(* IEC 61131-3 sources: nautilus/examples/lift-station/lib, 2 files *)

(* ---- physics.st ---- *)
(* Bench-only plant model: a wet-well level integrator and a submersible
   pump/VFD dynamic model. Two FUNCTION_BLOCKs, no PROGRAM — a project
   library (docs/functions.md "A .ld library", the same rule for .st).
   sim.st is the only caller; field.yaml has no sim task, so these two
   blocks sit compiled but unused in that manifest — harmless dead code,
   the same way a project's other library functions are. *)

FUNCTION_BLOCK WetWellModel
(* Integrates a level from an inflow/outflow balance. WW-101: a 13 ft
   level span over 1,320 gal of usable volume between the span's limits,
   so 13.2 gal per %: 100 gpm net moves the level 1 % in about 8 s. *)
VAR_INPUT
    InflowGpm  : REAL;
    OutflowGpm : REAL;
    Dt         : REAL; (* seconds *)
END_VAR
VAR_IN_OUT
    Level : REAL; (* %, 0..100 *)
END_VAR
VAR CONSTANT
    GalPerPercent : REAL := 13.2; (* 1,320 gal span / 100 % = 13.2 gal per % *)
END_VAR
(* gal/min * s / 60 = gal *)
Level := LIMIT(0.0, Level + (InflowGpm - OutflowGpm) * Dt / 60.0 / GalPerPercent, 100.0);
END_FUNCTION_BLOCK

FUNCTION_BLOCK VfdModel
(* A submersible pump + VFD, standing in for the field device on the
   bench: RunCmd/SpeedCmd in, Running/SpeedHz/Amps/Fault out. Running lags
   RunCmd by 0.5 s (starter contactor + soft-start), and drops the instant
   a fault is injected. SpeedHz ramps toward SpeedCmd at 10 Hz/s while
   commanded and running, and ramps back to 0 otherwise. Amps follows
   speed-squared, the affinity-law shape a centrifugal load actually
   draws. Fault is a plain pass-through of the bench inject tag — a real
   VFD's own fault relay, not the ladder's fail-to-run latch (that is a
   separate, higher-level condition computed in permissives.ld). *)
VAR_INPUT
    RunCmd      : BOOL;
    SpeedCmd    : REAL;
    Dt          : REAL;
    InjectFault : BOOL;
END_VAR
VAR_OUTPUT
    Running : BOOL;
    SpeedHz : REAL;
    Amps    : REAL;
    Fault   : BOOL;
END_VAR
VAR
    t1 : TON;
END_VAR
VAR CONSTANT
    RampHzPerS : REAL := 10.0; (* speed ramp rate *)
    FullLoadA  : REAL := 22.0; (* amps at MaxHz, full load *)
    MaxHz      : REAL := 60.0; (* VFD speed ceiling *)
END_VAR
Fault := InjectFault;
t1(IN := RunCmd AND NOT Fault, PT := T#500MS);
Running := t1.Q;
IF Running THEN
    SpeedHz := LIMIT(0.0, SpeedHz + LIMIT(-RampHzPerS * Dt, SpeedCmd - SpeedHz, RampHzPerS * Dt), MaxHz);
ELSE
    SpeedHz := MAX(0.0, SpeedHz - RampHzPerS * Dt);
END_IF;
Amps := (SpeedHz / MaxHz) * (SpeedHz / MaxHz) * FullLoadA;
END_FUNCTION_BLOCK

(* ---- pump.st ---- *)
(* Runtime accounting shared by both pumps: a retained UDT (PumpStats) and
   a FUNCTION_BLOCK that updates it by reference, so neither the sequence
   nor the permissives ever touch accumulation math themselves. A .st file
   with no PROGRAM is a project library — see docs/functions.md "A .ld
   library" (the same rule, one language over). *)

TYPE
  PumpStats : STRUCT
    Starts     : INT;   (* start count *)
    Hours      : REAL;  (* run hours *)
    LastRunSec : REAL;  (* length of the most recently completed run *)
  END_STRUCT;
END_TYPE

FUNCTION_BLOCK RuntimeMeter
(* Counts a start on Running's rising edge, accumulates run hours while
   Running, and captures the length of the run that just ended. Bound to
   the UDT tag by VAR_IN_OUT so two calls (P101_Stats, P102_Stats) each
   read and write their own copy — see docs/functions.md "VAR_IN_OUT is a
   reference pin". *)
VAR_INPUT
    Running : BOOL;
    Dt      : REAL; (* seconds since the last call *)
END_VAR
VAR_IN_OUT
    Stats : PumpStats;
END_VAR
VAR
    edgeUp   : R_TRIG;
    edgeDown : F_TRIG;
    runSec   : REAL;
END_VAR
edgeUp(CLK := Running);
edgeDown(CLK := Running);
IF edgeUp.Q THEN
    Stats.Starts := Stats.Starts + 1;
    runSec := 0.0;
END_IF;
IF Running THEN
    Stats.Hours := Stats.Hours + Dt / 3600.0;
    runSec := runSec + Dt;
END_IF;
IF edgeDown.Q THEN
    Stats.LastRunSec := runSec;
END_IF;
END_FUNCTION_BLOCK

FUNCTION PumpFlowGpm : REAL
(* Discharge flow at a given VFD speed — a rough affinity curve pinned to
   two points: ~0 gpm below 25 Hz (not enough head to open the check
   valve), 400 gpm at 60 Hz, linear between. Shared by the bench sim
   (lib/physics.st) and anywhere logic wants an expected flow from a
   commanded speed. *)
VAR_INPUT
    SpeedHz : REAL;
END_VAR
IF SpeedHz <= 25.0 THEN
    PumpFlowGpm := 0.0;
ELSE
    PumpFlowGpm := (SpeedHz - 25.0) / (60.0 - 25.0) * 400.0;
END_IF;
END_FUNCTION
